(* IEC 61131-3 sources: PLCHaT-dataset/benchmark_mutated/237_FB_ColorLightControl/mutation_2/syntax_check, 1 file *)

(* ---- 237_FB_ColorLightControl.st.clean.st ---- *)
FUNCTION_BLOCK FB_ColorLightControl
VAR_INPUT
    controlButton : BOOL;
END_VAR
VAR_OUTPUT
    greenLight : BOOL;
    redLight : BOOL;
    yellowLight : BOOL;
END_VAR
VAR
    currentState : INT := 0;
END_VAR

IF controlButton THEN
    currentState := currentState + 1;
    IF currentState > 6 THEN
        currentState := 1;
    END_IF;
END_IF;

CASE currentState OF
    1:
        greenLight := TRUE;
        redLight := FALSE;
        yellowLight := FALSE;
    2:
        greenLight := FALSE;
        redLight := TRUE;
        yellowLight := FALSE;
    3:
        greenLight := FALSE;
        redLight := FALSE;
        yellowLight := TRUE;
    4:
        greenLight := TRUE;
        redLight := TRUE;
        yellowLight := TRUE;
    5:
        greenLight := FALSE;
        redLight := FALSE;
        yellowLight := FALSE;
END_CASE;

END_FUNCTION_BLOCK
